TYPE TcoAbbRW_Status_v_8_2_x :
STRUCT
	ActionDescription : STRING(100);	
	State:TcoAbbRW_State_v_8_2_x;


END_STRUCT
END_TYPE

(* stored: Version 1.1.0.1, ProductVersion 3.1.4024.12
   DUT TcoAbbRW_Status_v_8_2_x: Id {7b9b9e61-f425-486c-a8e5-115cd80c0dc7} *)
